Fanuc KAREL source: kc00014.KL

-- PROVISIONAL review KL for V770-1; original PC SHA256 ba4363355d5bae2bcde231139c7cd044bc7c6db3ea1e38319adb0d5a90bae23a
-- Incomplete behavior may be omitted. Consult companion uncertainty JSON. Do not deploy.
PROGRAM KC00014
%NOLOCKGROUP
BEGIN
  -- UNRESOLVED_PC offsets 5-15; opcodes 27,31,23
  -- UNRESOLVED_PC offsets 20-24; opcodes 7F
END KC00014
